(* IEC 61131-3 sources: JingjiangArm/moonboxpro_arm_8.4/Application/Application/任务列表/Main_Task/IO配置表_1/OuNuo, 7 files *)

(* ---- KS_AbsEncModule_IODeal_OuNuo.st ---- *)
(*@CES
Name=KS_AbsEncModule_IODeal_OuNuo
Type=FunctionBlock
TypeGuid=6f9dac99-8de1-4efc-8465-68ac443b7d08
Guid=443b5ecb-ab70-45c9-9c02-718bc4c5ad3b
HasDeclaration=True
HasImplementation=False
*)
{DECLARATION}
FUNCTION_BLOCK KS_AbsEncModule_IODeal_OuNuo
VAR_INPUT
	i_xInputEn:BOOL;
	i_xOutPutEn:BOOL;
	(*这些值的处理未考虑双收双放*)
	i_pdwAbsEncSinglePos_Uw:POINTER TO DWORD;
	i_pwAbsEncMultiPos_Uw:POINTER TO WORD;
	(*收料*)
	i_pdwAbsEncSinglePos_Rw:POINTER TO DWORD;
	i_pwAbsEncMultiPos_Rw:POINTER TO WORD;
	//2025.08.20.152113+
	i_pstStAbsEncIOModule_Uw:POINTER TO StAbsEncIOModule;
	i_pstStAbsEncIOModule_Rw:POINTER TO StAbsEncIOModule;

END_VAR
VAR
	wIWTest:WORD;
	wQWTest: WORD;
	byAbsEncSts: BOOL;
END_VAR

{IMPLEMENTATION}

(* ---- KS_FB_IOMAP_AIAO_OuNuo.st ---- *)
(*@CES
Name=KS_FB_IOMAP_AIAO_OuNuo
Type=FunctionBlock
TypeGuid=6f9dac99-8de1-4efc-8465-68ac443b7d08
Guid=779e4782-a341-46a3-85b1-e10599855110
HasDeclaration=True
HasImplementation=False
*)
{DECLARATION}
FUNCTION_BLOCK KS_FB_IOMAP_AIAO_OuNuo
VAR_INPUT
	i_xEn: BOOL;(*功能块使能|*)
	i_xRdInput: BOOL;(*读io输入|*)
	i_xWrOutput: BOOL;(*写io输出|*)
	i_pstStSysParam								: POINTER TO StSysParam;
	i_pastStProgMonitoring						: POINTER TO ARRAY [1..2] OF StProgMonitoring;
END_VAR
VAR_OUTPUT
	o_xEno: BOOL;(*indicated to i_xEn|*)
	o_iErNo: INT;(*0.no err\-1.bad parameter|*)
END_VAR
VAR
	fb_KS_FB_SetAIType: KS_FB_SetAIType;
	fbKS_FB_Analog_IO_CTL: KS_FB_Analog_IO_CTL;

	byAiFilterTms_UwRw_I					:  BYTE:= 1;(*滤波次数*)
	byAiFilterTms_UwRw_II					:  BYTE:= 1;
	byAiFilterTms_IfOf_I					:  BYTE:= 1;
	byAiFilterTms_IfOf_II					:  BYTE:= 1;
	byAiFilterTms_DiaMeasure_I				:   BYTE:= 1;
	byAiFilterTms_DiaMeasure_II				:   BYTE:= 1;
END_VAR

{IMPLEMENTATION}

(* ---- KS_FB_IOMAP_Axis_OuNuo.st ---- *)
(*@CES
Name=KS_FB_IOMAP_Axis_OuNuo
Type=FunctionBlock
TypeGuid=6f9dac99-8de1-4efc-8465-68ac443b7d08
Guid=1c96003f-84aa-4353-ab1a-d2c99d7a7d11
HasDeclaration=True
HasImplementation=False
*)
{DECLARATION}
FUNCTION_BLOCK KS_FB_IOMAP_Axis_OuNuo
VAR_INPUT
	i_xEn: BOOL;(*功能块使能|*)
	i_xRdInput: BOOL;(*读io输入|*)
	i_xWrOutput: BOOL;(*写io输出|*)
	i_pastStIOMap_Axis_FE						: POINTER TO ARRAY [1..MAX_UNIT_NUM] OF StIOMap_Axis_FE;(*轴io数据区域|*)
END_VAR
VAR_OUTPUT
	o_xEno										: BOOL;(*indicated to i_xEn|*)
	o_iErNo										: INT;(*0.no err\-1.bad parameter|*)
END_VAR
VAR
	afbKS_FB_IOMap_Axis							: ARRAY [1..MAX_UNIT_NUM] OF KS_FB_MapAxisIOBasic;(*色组IO配置*)
END_VAR

{IMPLEMENTATION}

(* ---- KS_FB_IOMAP_AxisExtra_OuNuo.st ---- *)
(*@CES
Name=KS_FB_IOMAP_AxisExtra_OuNuo
Type=FunctionBlock
TypeGuid=6f9dac99-8de1-4efc-8465-68ac443b7d08
Guid=c18c8725-8f70-4642-a4b0-543efd8272e5
HasDeclaration=True
HasImplementation=False
*)
{DECLARATION}
FUNCTION_BLOCK KS_FB_IOMAP_AxisExtra_OuNuo
VAR_INPUT
	i_xEn: BOOL;(*功能块使能|*)
	i_xRdInput: BOOL;(*读io输入|*)
	i_xWrOutput: BOOL;(*写io输出|*)
	i_pastStIOMap_Axis_Extra_FE						: POINTER TO ARRAY [1..MAX_UNIT_NUM] OF StIOMap_Axis_Extra_FE;(*轴io数据区域|*)
	i_pstStSysParam	:POINTER TO StSysParam;
END_VAR
VAR_OUTPUT
	o_xEno										: BOOL;(*indicated to i_xEn|*)
	o_iErNo										: INT;(*0.no err\-1.bad parameter|*)
END_VAR
VAR
	afbKS_FB_IOMap_AxisExtra							: ARRAY [1..MAX_UNIT_NUM] OF KS_FB_MapAxisIOExtra;(*色组IO配置*)
END_VAR

{IMPLEMENTATION}

(* ---- KS_FB_IOMAP_Main_OuNuo.st ---- *)
(*@CES
Name=KS_FB_IOMAP_Main_OuNuo
Type=FunctionBlock
TypeGuid=6f9dac99-8de1-4efc-8465-68ac443b7d08
Guid=cafe5f1e-5342-4aa3-b5fa-17df2ef97cab
HasDeclaration=True
HasImplementation=False
*)
{DECLARATION}
FUNCTION_BLOCK KS_FB_IOMAP_Main_OuNuo
(*主面板IO配置分A/B系和放/收牵*)
(*正常单收单放选1和2*)
(*双收双放1和2是A系的放牵收牵，3和4是B系的放牵收牵*)
(*双收双放A放B收1和4*)
VAR_INPUT
	i_xEn: BOOL;(*功能块使能|*)
	i_xRdInput: BOOL;(*读io输入|*)
	i_xWrOutput: BOOL;(*写io输出|*)
	i_pastStIOMap_Main_FE						: POINTER TO ARRAY [1..4] OF StIOMap_Main_FE;(*轴io数据区域|*)
END_VAR
VAR_OUTPUT
	o_xEno										: BOOL;(*indicated to i_xEn|*)
	o_iErNo										: INT;(*0.no err\-1.bad parameter|*)
END_VAR
VAR
	afbKS_FB_MapIO_Main						: ARRAY [1..4] OF KS_FB_MapIO_Main;(*主面板IO配置*)
END_VAR

{IMPLEMENTATION}

(* ---- KS_FB_IOMAP_UwRw_OuNuo.st ---- *)
(*@CES
Name=KS_FB_IOMAP_UwRw_OuNuo
Type=FunctionBlock
TypeGuid=6f9dac99-8de1-4efc-8465-68ac443b7d08
Guid=cd72dcdb-6cfc-465e-91fc-8c9132cffc39
HasDeclaration=True
HasImplementation=False
*)
{DECLARATION}
 FUNCTION_BLOCK KS_FB_IOMAP_UwRw_OuNuo
VAR_INPUT
	i_xEn: BOOL;(*功能块使能|*)
	i_xRdInput: BOOL;(*读io输入|*)
	i_xWrOutput: BOOL;(*写io输出|*)
	i_pastStIOMap_UwRw_FE_Uw					: POINTER TO ARRAY [1..2] OF StIOMap_UwRw_FE;(*轴io数据区域|*)
	i_pastStIOMap_UwRw_FE_Rw					: POINTER TO ARRAY [1..2] OF StIOMap_UwRw_FE;(*轴io数据区域|*)
END_VAR
VAR_OUTPUT
	o_xEno										: BOOL;(*indicated to i_xEn|*)
	o_iErNo										: INT;(*0.no err\-1.bad parameter|*)
END_VAR
VAR
	afbKS_FB_MapIO_UwRw_Uw						: ARRAY [1..2] OF KS_FB_MapIO_UwRw;
	afbKS_FB_MapIO_UwRw_Rw						: ARRAY [1..2] OF KS_FB_MapIO_UwRw;
END_VAR

{IMPLEMENTATION}

(* ---- KS_FB_StepDriveIODeal_OuNuo.st ---- *)
(*@CES
Name=KS_FB_StepDriveIODeal_OuNuo
Type=FunctionBlock
TypeGuid=6f9dac99-8de1-4efc-8465-68ac443b7d08
Guid=968bd9c6-1e80-4b52-be82-587a9a1cb845
HasDeclaration=True
HasImplementation=False
*)
{DECLARATION}
FUNCTION_BLOCK KS_FB_StepDriveIODeal_OuNuo
VAR_INPUT
	i_xInputEn:BOOL;
	i_xOutPutEn:BOOL;
	i_pastStDigitalMicroStepDrive :POINTER TO  ARRAY [1..MAX_UNIT_NUM] OF StDigitalMicroStepDrive;
	i_pastStStepDriveIOModule:POINTER TO ARRAY [1..MAX_UNIT_NUM] OF StStepDriveIOModule;
	i_pastStEnc0410R:POINTER TO ARRAY [1..MAX_UNIT_NUM] OF StEnc0410R;
END_VAR
VAR_OUTPUT
END_VAR
VAR
	wTest: WORD;
	afbKS_FB_StepDriveIOModule: ARRAY [1..MAX_UNIT_NUM] OF KS_FB_StepDriveIOModule;
END_VAR

{IMPLEMENTATION}
